Staubli VAL3: isPointOK.pgx

public program isPointOK(string x_sKey, num x_nIndex, bool& x_bResult)
  local pointRx l_pPoint
  local num l_nToolID
  local tool l_tTool
  local frame l_fFrame
  local num l_nFrameID
  local bool l_bResult
  local jointRx l_jResult
begin
  link(l_tTool,flange)
  link(l_fFrame,world)
  call getFrameID(x_sKey,l_nFrameID)
  call getToolID(x_sKey,l_nToolID)
  call savedata:getTool(l_nToolID,l_tTool)
  call savedata:getFrame(l_nFrameID,l_fFrame)
  link(l_pPoint,l_fFrame)
  l_pPoint.trsf=trajTemp:tTrajItem[x_sKey].pPointItem[x_nIndex].pPointRx.trsf
  l_pPoint.config=trajTemp:tTrajItem[x_sKey].pPointItem[x_nIndex].pPointRx.config

  l_bResult=pointToJoint(l_tTool,herej(),l_pPoint,l_jResult)
  if l_pPoint.trsf!={0,0,0,0,0,0} and l_bResult and isInRange(l_jResult)
    x_bResult=true
  else
    x_bResult=false
  endIf
end
